// TwinCAT 3 PLC project PlcKessel
// Title: PlcKessel
// project tree:
//   DUTs/ E_Zustand.TcDUT
//   POUs/ I_Maschine.TcPOU, FB_Maschine.TcPOU, FB_Kessel.TcPOU, MAIN.TcPOU
//   GVLs/ GVL.TcGVL

// ---- DUTs/E_Zustand.TcDUT
TYPE E_Zustand :
(
	Aus := 0,
	Bereit := 1,
	Heizen := 2,
	Warnung := 3,
	Kritisch := 4,
	Notaus := 5
);
END_TYPE

// ---- GVLs/GVL.TcGVL
{attribute 'qualified_only'}
VAR_GLOBAL
	// Komutlar (ADS schreibt, FB_Kessel verarbeitet)
	CmdHeizung : BOOL;
	CmdPumpe : BOOL := TRUE;
	CmdSollwert : LREAL := 60.0;
	CmdNotaus : BOOL;
	CmdNotausReset : BOOL;

	// Zustand (ADS liest, nur PLC schreibt)
	Temperatur : LREAL := 20.0;
	Heizung : BOOL;
	Pumpe : BOOL := TRUE;
	Sollwert : LREAL := 60.0;
	Notaus : BOOL;
	ZielAlarmSekunden : LREAL;
	AutoGestoppt : BOOL;
END_VAR

// ---- POUs/FB_Kessel.TcPOU
FUNCTION_BLOCK FB_Kessel EXTENDS FB_Maschine
VAR CONSTANT
	WarnSchwelle : LREAL := 80.0;
	KritischSchwelle : LREAL := 90.0;
	UmgebungsTemperatur : LREAL := 20.0;
	HeizrateProSekunde : LREAL := 0.5;
	KuehlrateProSekunde : LREAL := 0.25;
	Jitter : LREAL := 0.3;
	Hysterese : LREAL := 0.5;
END_VAR
VAR
	_temperatur : LREAL := 20.0;
	_heizung : BOOL;
	_pumpe : BOOL := TRUE;
	_sollwert : LREAL := 60.0;
	_zielAlarmSekunden : LREAL;
	_autoGestoppt : BOOL;
	_automatik : BOOL := TRUE;
	_zufallSeed : UDINT := 12345;
	_gestartet : BOOL;
	_cmdHeizungAlt : BOOL;
	_cmdPumpeAlt : BOOL := TRUE;
	_cmdSollwertAlt : LREAL := 60.0;
END_VAR

// Einmaliger Selbststart beim ersten Zyklus (Start/Stop bleiben als OOP-Methoden verfügbar).
IF NOT _gestartet THEN
	Start();
	_gestartet := TRUE;
END_IF

VerarbeiteBefehle();
Aktualisiere(0.1);
SchreibeZustand();

METHOD NotausAusloesen
SUPER^.NotausAusloesen();
_heizung := FALSE;
_pumpe := FALSE;
_zielAlarmSekunden := 0.0;
END_METHOD

METHOD NotausZuruecksetzen
SUPER^.NotausZuruecksetzen();
_automatik := TRUE;
_autoGestoppt := FALSE;
_zielAlarmSekunden := 0.0;
END_METHOD

METHOD PRIVATE VerarbeiteBefehle
// Notaus / Reset werden als Impuls konsumiert.
IF GVL.CmdNotaus THEN
	NotausAusloesen();
	GVL.CmdNotaus := FALSE;
END_IF

IF GVL.CmdNotausReset THEN
	NotausZuruecksetzen();
	GVL.CmdNotausReset := FALSE;
END_IF

// Alle anderen Befehle nur, wenn nicht verriegelt.
IF NOT _notaus THEN
	// Sollwert (Pegel, mit Klemmung 0..100 °C)
	IF GVL.CmdSollwert <> _cmdSollwertAlt THEN
		_cmdSollwertAlt := GVL.CmdSollwert;
		_sollwert := LIMIT(0.0, GVL.CmdSollwert, 100.0);
		_autoGestoppt := FALSE;
	END_IF

	// Heizung (manuell, Flanke)
	IF GVL.CmdHeizung <> _cmdHeizungAlt THEN
		_cmdHeizungAlt := GVL.CmdHeizung;
		_heizung := GVL.CmdHeizung;
		_automatik := FALSE;
		IF GVL.CmdHeizung THEN
			_autoGestoppt := FALSE;
		END_IF
	END_IF

	// Pumpe (manuell, Flanke)
	IF GVL.CmdPumpe <> _cmdPumpeAlt THEN
		_cmdPumpeAlt := GVL.CmdPumpe;
		_pumpe := GVL.CmdPumpe;
	END_IF
END_IF
END_METHOD

METHOD PRIVATE Aktualisiere
VAR_INPUT
	sekunden : LREAL;
END_VAR
IF _zustand = E_Zustand.Aus THEN
	RETURN;
END_IF

sekunden := LIMIT(0.0, sekunden, 1.0);

IF _notaus THEN
	_heizung := FALSE;
	_pumpe := FALSE;
	_zielAlarmSekunden := 0.0;
	_temperatur := Annaehern(_temperatur, UmgebungsTemperatur, KuehlrateProSekunde * sekunden);
ELSE
	IF _automatik THEN
		IF _heizung AND (_temperatur >= _sollwert + Hysterese) THEN
			_heizung := FALSE;
		ELSIF (NOT _heizung) AND (_temperatur < _sollwert - Hysterese) THEN
			_heizung := TRUE;
		END_IF
	END_IF

	IF _heizung THEN
		_temperatur := _temperatur + HeizrateProSekunde * sekunden;
	ELSE
		_temperatur := Annaehern(_temperatur, UmgebungsTemperatur, KuehlrateProSekunde * sekunden);
	END_IF

	// Kritisch: ab 90 °C wird die Heizung automatisch abgeschaltet.
	IF _temperatur >= KritischSchwelle THEN
		_heizung := FALSE;
	END_IF

	// Ziel erreicht: Alarm + Countdown, danach automatische Abschaltung.
	IF _heizung AND (_temperatur >= _sollwert) AND (_zielAlarmSekunden <= 0.0) THEN
		_zielAlarmSekunden := 5.0;
	END_IF

	IF _zielAlarmSekunden > 0.0 THEN
		IF (NOT _automatik) AND (NOT _heizung) THEN
			_zielAlarmSekunden := 0.0;
		ELSE
			_zielAlarmSekunden := _zielAlarmSekunden - sekunden;
			IF _zielAlarmSekunden <= 0.0 THEN
				_zielAlarmSekunden := 0.0;
				_heizung := FALSE;
				_automatik := FALSE;
				_autoGestoppt := TRUE;
			END_IF
		END_IF
	END_IF
END_IF

// Rauschanteil (±Jitter) und Grenzbereich.
_temperatur := _temperatur + Zufall() * Jitter * sekunden;
_temperatur := LIMIT(10.0, _temperatur, 120.0);

// Zustand ableiten.
IF _notaus THEN
	_zustand := E_Zustand.Notaus;
ELSIF _temperatur >= KritischSchwelle THEN
	_zustand := E_Zustand.Kritisch;
ELSIF _temperatur >= WarnSchwelle THEN
	_zustand := E_Zustand.Warnung;
ELSIF _heizung THEN
	_zustand := E_Zustand.Heizen;
ELSE
	_zustand := E_Zustand.Bereit;
END_IF
END_METHOD

METHOD PRIVATE SchreibeZustand
// Durum değişkenleri yalnızca PLC tarafından yazılır; ADS sadece okur.
GVL.Temperatur := _temperatur;
GVL.Heizung := _heizung;
GVL.Pumpe := _pumpe;
GVL.Sollwert := _sollwert;
GVL.Notaus := _notaus;
GVL.ZielAlarmSekunden := _zielAlarmSekunden;
GVL.AutoGestoppt := _autoGestoppt;
END_METHOD

METHOD PRIVATE Annaehern : LREAL
VAR_INPUT
	aktuell : LREAL;
	ziel : LREAL;
	schritt : LREAL;
END_VAR
IF aktuell < ziel THEN
	Annaehern := MIN(ziel, aktuell + schritt);
ELSIF aktuell > ziel THEN
	Annaehern := MAX(ziel, aktuell - schritt);
ELSE
	Annaehern := aktuell;
END_IF
END_METHOD

METHOD PRIVATE Zufall : LREAL
// Einfacher linearer Kongruenzgenerator: Wert in [-1, 1).
_zufallSeed := (_zufallSeed * 1664525) + 1013904223;
Zufall := (UDINT_TO_LREAL(_zufallSeed) / 2147483648.0) - 1.0;
END_METHOD

PROPERTY Temperatur : LREAL
END_PROPERTY

END_FUNCTION_BLOCK

// ---- POUs/FB_Maschine.TcPOU
FUNCTION_BLOCK FB_Maschine IMPLEMENTS I_Maschine
VAR
	_zustand : E_Zustand := E_Zustand.Aus;
	_notaus : BOOL := FALSE;
END_VAR

METHOD Start
IF NOT _notaus THEN
	_zustand := E_Zustand.Bereit;
END_IF
END_METHOD

METHOD Stop
_zustand := E_Zustand.Aus;
END_METHOD

METHOD NotausAusloesen
_notaus := TRUE;
_zustand := E_Zustand.Notaus;
END_METHOD

METHOD NotausZuruecksetzen
_notaus := FALSE;
_zustand := E_Zustand.Bereit;
END_METHOD

PROPERTY Zustand : E_Zustand
END_PROPERTY

END_FUNCTION_BLOCK

// ---- POUs/I_Maschine.TcPOU
INTERFACE I_Maschine

METHOD Start
END_METHOD

METHOD Stop
END_METHOD

METHOD NotausAusloesen
END_METHOD

METHOD NotausZuruecksetzen
END_METHOD

END_INTERFACE

// ---- POUs/MAIN.TcPOU
PROGRAM MAIN
VAR
	fbKessel : FB_Kessel;
END_VAR

// Ein Aufruf pro Task-Zyklus (Zykluszeit z. B. 100 ms).
fbKessel();

END_PROGRAM
